(* IEC 61131-3 sources: plc-st-coding-agent/progress/evidence/v13_rescore_20261108b/candidates/custom_deepseek-v4pro, 35 files *)

(* ---- public-easy-01.st ---- *)
FUNCTION_BLOCK FB
VAR_INPUT
    bottleSensor: BOOL;
    cleaningConfirmButton: BOOL;
    fillingConfirmButton: BOOL;
    cappingConfirmButton: BOOL;
    packingConfirmButton: BOOL;
    finishedButton: BOOL;
END_VAR
VAR_OUTPUT
    Pump_Motor: BOOL;
    Filling_Valve: BOOL;
    Capping_Machine: BOOL;
    Packing_Machine: BOOL;
    Completion_Light: BOOL;
END_VAR
VAR
    step: INT := 0;
END_VAR

IF finishedButton THEN
    step := 0;
    Pump_Motor := FALSE;
    Filling_Valve := FALSE;
    Capping_Machine := FALSE;
    Packing_Machine := FALSE;
    Completion_Light := FALSE;
ELSE
    CASE step OF
        0:
            IF bottleSensor THEN
                step := 1;
                Pump_Motor := TRUE;
                Filling_Valve := FALSE;
                Capping_Machine := FALSE;
                Packing_Machine := FALSE;
                Completion_Light := FALSE;
            ELSE
                Pump_Motor := FALSE;
                Filling_Valve := FALSE;
                Capping_Machine := FALSE;
                Packing_Machine := FALSE;
                Completion_Light := FALSE;
            END_IF

        1:
            Pump_Motor := TRUE;
            Filling_Valve := FALSE;
            Capping_Machine := FALSE;
            Packing_Machine := FALSE;
            Completion_Light := FALSE;
            IF cleaningConfirmButton THEN
                step := 2;
                Filling_Valve := TRUE;
            END_IF

        2:
            Pump_Motor := TRUE;
            Filling_Valve := TRUE;
            Capping_Machine := FALSE;
            Packing_Machine := FALSE;
            Completion_Light := FALSE;
            IF fillingConfirmButton THEN
                step := 3;
                Capping_Machine := TRUE;
            END_IF

        3:
            Pump_Motor := TRUE;
            Filling_Valve := TRUE;
            Capping_Machine := TRUE;
            Packing_Machine := FALSE;
            Completion_Light := FALSE;
            IF cappingConfirmButton THEN
                step := 4;
                Packing_Machine := TRUE;
            END_IF

        4:
            Pump_Motor := TRUE;
            Filling_Valve := TRUE;
            Capping_Machine := TRUE;
            Packing_Machine := TRUE;
            Completion_Light := FALSE;
            IF packingConfirmButton THEN
                step := 5;
                Completion_Light := TRUE;
            END_IF

        5:
            Pump_Motor := TRUE;
            Filling_Valve := TRUE;
            Capping_Machine := TRUE;
            Packing_Machine := TRUE;
            Completion_Light := TRUE;

    ELSE
        step := 0;
        Pump_Motor := FALSE;
        Filling_Valve := FALSE;
        Capping_Machine := FALSE;
        Packing_Machine := FALSE;
        Completion_Light := FALSE;
    END_CASE
END_IF

END_FUNCTION_BLOCK

(* ---- public-easy-02.st ---- *)
FUNCTION_BLOCK FB
VAR_INPUT
    value : DWORD;
END_VAR
VAR_OUTPUT
    hasChanged : BOOL;
    hasRisingEdges : BOOL;
    risingBits : DWORD;
    noOfRisingBits : USINT;
    hasFallingEdges : BOOL;
    fallingBits : DWORD;
    noOfFallingBits : USINT;
END_VAR
VAR
    previousValue : DWORD := 0;
    bitIndex : INT;
END_VAR
    risingBits := value AND (NOT previousValue);
    fallingBits := (NOT value) AND previousValue;

    hasRisingEdges := risingBits <> 0;
    hasFallingEdges := fallingBits <> 0;
    hasChanged := hasRisingEdges OR hasFallingEdges;

    noOfRisingBits := 0;
    noOfFallingBits := 0;
    FOR bitIndex := 0 TO 31 DO
        IF (risingBits AND SHL(DWORD#1, bitIndex)) <> 0 THEN
            noOfRisingBits := noOfRisingBits + 1;
        END_IF;
        IF (fallingBits AND SHL(DWORD#1, bitIndex)) <> 0 THEN
            noOfFallingBits := noOfFallingBits + 1;
        END_IF;
    END_FOR;

    previousValue := value;
END_FUNCTION_BLOCK

(* ---- public-easy-03.st ---- *)
FUNCTION_BLOCK FB
VAR_INPUT
    Value : REAL;
    hiLevel : REAL;
    loLevel : REAL;
    hystWindow : REAL;
END_VAR
VAR_OUTPUT
    hiAlarm : BOOL;
    loAlarm : BOOL;
    error : BOOL;
    status : WORD;
END_VAR
VAR
END_VAR

error := FALSE;
status := 0;

IF loLevel >= hiLevel THEN
    error := TRUE;
    status := 16#8001;
ELSIF hystWindow >= (hiLevel - loLevel) THEN
    error := TRUE;
    status := 16#8002;
ELSE
    IF Value > hiLevel THEN
        hiAlarm := TRUE;
    ELSIF Value < (hiLevel - hystWindow) THEN
        hiAlarm := FALSE;
    END_IF;

    IF Value < loLevel THEN
        loAlarm := TRUE;
    ELSIF Value > (loLevel + hystWindow) THEN
        loAlarm := FALSE;
    END_IF;
END_IF;

END_FUNCTION_BLOCK

(* ---- public-easy-04.st ---- *)
FUNCTION_BLOCK FB
VAR_INPUT
    VISCOSITY_OK: BOOL;
    PASTE_E_STOP_NC: BOOL;
    DebounceTime: TIME;
    CycleTime: TIME;
END_VAR
VAR_OUTPUT
    VFD_RUN: BOOL;
    PUMP_MAINT_DUE: BOOL;
    PUMP_RUNTIME_ACC: LINT;
END_VAR
VAR
    DebounceAccum: LINT := 0;               (* Debounce accumulated time in ms *)
    AccumRuntime: LINT := 0;                (* Accumulated pump runtime in ms *)
    MaintDue: BOOL := FALSE;                (* Maintenance due latch *)
    DebounceTimeMs: LINT := 0;              (* DebounceTime in ms *)
    MAINT_THRESHOLD: LINT := 1800000000;    (* 500 hours in ms *)
END_VAR

(* Convert DebounceTime to milliseconds (CODESYS TIME_TO_LINT preserves ms value) *)
DebounceTimeMs := TIME_TO_LINT(DebounceTime);

(* Debounce logic with E-stop priority:
   - VISCOSITY_OK FALSE immediately clears debounce.
   - E-stop active clears only incomplete debounce, keeps completed condition.
   - Normal condition accumulates when signal is stable and E-stop is OK.
*)
IF NOT VISCOSITY_OK THEN
    DebounceAccum := 0;
ELSIF NOT PASTE_E_STOP_NC THEN
    IF DebounceAccum < DebounceTimeMs THEN
        DebounceAccum := 0;
    END_IF;
ELSE
    IF DebounceAccum < DebounceTimeMs THEN
        DebounceAccum := DebounceAccum + TIME_TO_LINT(CycleTime);
        IF DebounceAccum > DebounceTimeMs THEN
            DebounceAccum := DebounceTimeMs;
        END_IF;
    END_IF;
END_IF;

(* Run command requires E-stop OK, viscosity raw signal TRUE and debounced condition valid *)
VFD_RUN := PASTE_E_STOP_NC AND VISCOSITY_OK AND (DebounceAccum >= DebounceTimeMs);

(* Accumulate enabled runtime only while pump is running *)
IF VFD_RUN THEN
    AccumRuntime := AccumRuntime + TIME_TO_LINT(CycleTime);
END_IF;

(* Maintenance due latch when accumulated time reaches 500 hours (1,800,000,000 ms) *)
IF AccumRuntime >= MAINT_THRESHOLD THEN
    MaintDue := TRUE;
END_IF;

(* Map internal state to outputs *)
PUMP_RUNTIME_ACC := AccumRuntime;
PUMP_MAINT_DUE := MaintDue;

END_FUNCTION_BLOCK

(* ---- public-easy-05.st ---- *)
FUNCTION_BLOCK FB
VAR_INPUT
    Gap_Exceeded : BOOL;
    Weld_E_Stop_NC : BOOL;
    DebounceTime : TIME;
END_VAR
VAR_OUTPUT
    Operator_Alert : BOOL;
    Weld_Soft_Start_Active : BOOL;
END_VAR
VAR
    init_count : DINT := 0;
    debounce_count : DINT := 0;
    InitPeriods : DINT := 5;
    DebouncePeriods : DINT;
END_VAR

DebouncePeriods := TIME_TO_DINT(DebounceTime);
IF DebouncePeriods < 3 THEN
    DebouncePeriods := 3;
END_IF;

Weld_Soft_Start_Active := (init_count < InitPeriods);

IF init_count < InitPeriods THEN
    init_count := init_count + 1;
END_IF;

IF NOT Weld_E_Stop_NC THEN
    Operator_Alert := FALSE;
    debounce_count := 0;
ELSE
    IF Weld_Soft_Start_Active THEN
        Operator_Alert := FALSE;
        debounce_count := 0;
    ELSE
        IF Gap_Exceeded THEN
            IF debounce_count < DebouncePeriods THEN
                debounce_count := debounce_count + 1;
            END_IF;
            IF debounce_count >= DebouncePeriods THEN
                Operator_Alert := TRUE;
            ELSE
                Operator_Alert := FALSE;
            END_IF;
        ELSE
            debounce_count := 0;
            Operator_Alert := FALSE;
        END_IF;
    END_IF;
END_IF;

END_FUNCTION_BLOCK

(* ---- public-easy-06.st ---- *)
FUNCTION_BLOCK FB
VAR_INPUT
    DO_LOW : BOOL;
    AERATION_E_STOP_NC : BOOL;
END_VAR
VAR_OUTPUT
    BLOWER_RUN : BOOL;
    AERATION_BLOWER_CYCLE_COUNT : UINT;
END_VAR
VAR
    timer_count : UINT := 0;
    last_run : BOOL := FALSE;
    run_cmd : BOOL := FALSE;
    cycle_count : UINT := 0;
END_VAR

IF DO_LOW AND AERATION_E_STOP_NC THEN
    IF timer_count < 5 THEN
        timer_count := timer_count + 1;
    END_IF;
ELSE
    timer_count := 0;
END_IF;

run_cmd := DO_LOW AND AERATION_E_STOP_NC AND (timer_count >= 5);

IF run_cmd AND NOT last_run THEN
    cycle_count := cycle_count + 1;
END_IF;

BLOWER_RUN := run_cmd;
AERATION_BLOWER_CYCLE_COUNT := cycle_count;
last_run := run_cmd;

END_FUNCTION_BLOCK

(* ---- public-hard-01.st ---- *)
FUNCTION_BLOCK FB
VAR_INPUT
    estop : BOOL;
    opeMode : BOOL;
    valveAStart : BOOL;
    valveBStart : BOOL;
    valveCStart : BOOL;
    valveDStart : BOOL;
    mixMotorStart : BOOL;
    autoStart : BOOL;
    processMode : BOOL;
    levelSensor : INT;
    mixMotorComplete : BOOL;
END_VAR
VAR_OUTPUT
    valveARun : BOOL;
    valveBRun : BOOL;
    valveCRun : BOOL;
    valveDRun : BOOL;
    mixMotorRun : BOOL;
END_VAR
VAR
    manValveA : BOOL := FALSE;
    manValveB : BOOL := FALSE;
    manValveC : BOOL := FALSE;
    manValveD : BOOL := FALSE;
    manMixMotor : BOOL := FALSE;
    autoStep : INT := 0;
    autoValveA : BOOL := FALSE;
    autoValveB : BOOL := FALSE;
    autoValveC : BOOL := FALSE;
    autoValveD : BOOL := FALSE;
    autoMixMotor : BOOL := FALSE;
    lastValveAStart : BOOL := FALSE;
    lastValveBStart : BOOL := FALSE;
    lastValveCStart : BOOL := FALSE;
    lastValveDStart : BOOL := FALSE;
    lastMixMotorStart : BOOL := FALSE;
    lastAutoStart : BOOL := FALSE;
    lastMixMotorComplete : BOOL := FALSE;
    lastOpeMode : BOOL := FALSE;
    valveAStartRising : BOOL;
    valveBStartRising : BOOL;
    valveCStartRising : BOOL;
    valveDStartRising : BOOL;
    mixMotorStartRising : BOOL;
    autoStartRising : BOOL;
    mixMotorCompleteRising : BOOL;
END_VAR

// 计算所有输入信号的上升沿
valveAStartRising := valveAStart AND NOT lastValveAStart;
valveBStartRising := valveBStart AND NOT lastValveBStart;
valveCStartRising := valveCStart AND NOT lastValveCStart;
valveDStartRising := valveDStart AND NOT lastValveDStart;
mixMotorStartRising := mixMotorStart AND NOT lastMixMotorStart;
autoStartRising := autoStart AND NOT lastAutoStart;
mixMotorCompleteRising := mixMotorComplete AND NOT lastMixMotorComplete;

// 急停或模式切换时，复位所有内部状态（手动记忆和自动步序）
IF (estop = FALSE) OR (opeMode <> lastOpeMode) THEN
    manValveA := FALSE;
    manValveB := FALSE;
    manValveC := FALSE;
    manValveD := FALSE;
    manMixMotor := FALSE;
    autoStep := 0;
    autoValveA := FALSE;
    autoValveB := FALSE;
    autoValveC := FALSE;
    autoValveD := FALSE;
    autoMixMotor := FALSE;
END_IF;

// 根据急停和模式设置输出
IF estop = TRUE THEN
    IF opeMode = FALSE THEN
        // 手动模式：按钮上升沿翻转对应输出
        IF valveAStartRising THEN
            manValveA := NOT manValveA;
        END_IF;
        IF valveBStartRising THEN
            manValveB := NOT manValveB;
        END_IF;
        IF valveCStartRising THEN
            manValveC := NOT manValveC;
        END_IF;
        IF valveDStartRising THEN
            manValveD := NOT manValveD;
        END_IF;
        IF mixMotorStartRising THEN
            manMixMotor := NOT manMixMotor;
        END_IF;

        valveARun := manValveA;
        valveBRun := manValveB;
        valveCRun := manValveC;
        valveDRun := manValveD;
        mixMotorRun := manMixMotor;
    ELSE
        // 自动模式
        IF autoStartRising THEN
            autoStep := 1;  // 进入FILL_A
            autoValveA := TRUE;
            autoValveB := FALSE;
            autoValveC := FALSE;
            autoValveD := FALSE;
            autoMixMotor := FALSE;
        END_IF;

        CASE autoStep OF
            0: // 空闲
                autoValveA := FALSE;
                autoValveB := FALSE;
                autoValveC := FALSE;
                autoValveD := FALSE;
                autoMixMotor := FALSE;

            1: // 填充A
                autoValveA := TRUE;
                autoValveB := FALSE;
                autoValveC := FALSE;
                autoValveD := FALSE;
                autoMixMotor := FALSE;
                IF levelSensor >= 50 THEN
                    autoValveA := FALSE;
                    autoStep := 2;
                END_IF;

            2: // 填充B
                autoValveB := TRUE;
                autoValveA := FALSE;
                autoValveC := FALSE;
                autoValveD := FALSE;
                autoMixMotor := FALSE;
                IF levelSensor >= 80 THEN
                    autoValveB := FALSE;
                    IF processMode THEN
                        autoStep := 4; // 填充C
                    ELSE
                        autoStep := 3; // 混合
                    END_IF;
                END_IF;

            3: // 混合电机运行
                autoMixMotor := TRUE;
                autoValveA := FALSE;
                autoValveB := FALSE;
                autoValveC := FALSE;
                autoValveD := FALSE;
                IF mixMotorCompleteRising THEN
                    autoMixMotor := FALSE;
                    autoValveD := TRUE;
                    autoStep := 5; // 出料
                END_IF;

            4: // 填充C（仅processMode=TRUE）
                autoValveC := TRUE;
                autoValveA := FALSE;
                autoValveB := FALSE;
                autoValveD := FALSE;
                autoMixMotor := FALSE;
                IF levelSensor >= 100 THEN
                    autoValveC := FALSE;
                    autoStep := 3; // 混合
                END_IF;

            5: // 出料
                autoValveD := TRUE;
                autoValveA := FALSE;
                autoValveB := FALSE;
                autoValveC := FALSE;
                autoMixMotor := FALSE;
                // 等待新的autoStart上升沿，由外层处理

            ELSE
                // 非法状态，复位
                autoStep := 0;
                autoValveA := FALSE;
                autoValveB := FALSE;
                autoValveC := FALSE;
                autoValveD := FALSE;
                autoMixMotor := FALSE;
        END_CASE;

        valveARun := autoValveA;
        valveBRun := autoValveB;
        valveCRun := autoValveC;
        valveDRun := autoValveD;
        mixMotorRun := autoMixMotor;
    END_IF;
ELSE
    // 急停触发：所有输出停止
    valveARun := FALSE;
    valveBRun := FALSE;
    valveCRun := FALSE;
    valveDRun := FALSE;
    mixMotorRun := FALSE;
END_IF;

// 更新历史值
lastValveAStart := valveAStart;
lastValveBStart := valveBStart;
lastValveCStart := valveCStart;
lastValveDStart := valveDStart;
lastMixMotorStart := mixMotorStart;
lastAutoStart := autoStart;
lastMixMotorComplete := mixMotorComplete;
lastOpeMode := opeMode;

END_FUNCTION_BLOCK

(* ---- public-hard-02.st ---- *)
FUNCTION_BLOCK FB
VAR_INPUT
    processLength : USINT;
    sensor1 : BOOL;
    sensor2 : BOOL;
    sensor3 : BOOL;
    sensor4 : BOOL;
    sensor5 : BOOL;
    station1Start : BOOL;
    station2Complete : BOOL;
    station3Complete : BOOL;
    station4Complete : BOOL;
    processSequence : ARRAY[1..8] OF USINT;
END_VAR
VAR_OUTPUT
    conveyorLeft : BOOL;
    conveyorRight : BOOL;
END_VAR
VAR
    phase : USINT := 0;
    curStation : USINT := 1;
    idx : USINT := 1;
    dstStation : USINT := 0;
    station1StartPrev : BOOL := FALSE;
    station2CompletePrev : BOOL := FALSE;
    station3CompletePrev : BOOL := FALSE;
    station4CompletePrev : BOOL := FALSE;
    sensor2Prev : BOOL := FALSE;
    sensor3Prev : BOOL := FALSE;
    sensor4Prev : BOOL := FALSE;
    sensor5Prev : BOOL := FALSE;
    station1StartRising : BOOL;
    station2CompleteRising : BOOL;
    station3CompleteRising : BOOL;
    station4CompleteRising : BOOL;
    sensor2Rising : BOOL;
    sensor3Rising : BOOL;
    sensor4Rising : BOOL;
    sensor5Rising : BOOL;
END_VAR

    station1StartRising := station1Start AND NOT station1StartPrev;
    station2CompleteRising := station2Complete AND NOT station2CompletePrev;
    station3CompleteRising := station3Complete AND NOT station3CompletePrev;
    station4CompleteRising := station4Complete AND NOT station4CompletePrev;
    sensor2Rising := sensor2 AND NOT sensor2Prev;
    sensor3Rising := sensor3 AND NOT sensor3Prev;
    sensor4Rising := sensor4 AND NOT sensor4Prev;
    sensor5Rising := sensor5 AND NOT sensor5Prev;

    IF phase = 0 THEN
        IF station1StartRising AND sensor1 THEN
            curStation := 1;
            idx := 1;
            dstStation := processSequence[idx];
            phase := 1;
        END_IF;
    ELSIF phase = 1 THEN
        IF (dstStation = 2 AND sensor2Rising) OR
           (dstStation = 3 AND sensor3Rising) OR
           (dstStation = 4 AND sensor4Rising) OR
           (dstStation = 5 AND sensor5Rising) THEN
            curStation := dstStation;
            IF dstStation = 5 THEN
                phase := 0;
                idx := 0;
            ELSE
                phase := 2;
            END_IF;
        END_IF;
    ELSIF phase = 2 THEN
        IF (curStation = 2 AND station2CompleteRising) OR
           (curStation = 3 AND station3CompleteRising) OR
           (curStation = 4 AND station4CompleteRising) THEN
            idx := idx + 1;
            dstStation := processSequence[idx];
            phase := 1;
        END_IF;
    ELSE
        phase := 0;
    END_IF;

    IF phase = 1 THEN
        IF dstStation > curStation THEN
            conveyorRight := TRUE;
            conveyorLeft := FALSE;
        ELSIF dstStation < curStation THEN
            conveyorLeft := TRUE;
            conveyorRight := FALSE;
        ELSE
            conveyorLeft := FALSE;
            conveyorRight := FALSE;
        END_IF;
    ELSE
        conveyorLeft := FALSE;
        conveyorRight := FALSE;
    END_IF;

    station1StartPrev := station1Start;
    station2CompletePrev := station2Complete;
    station3CompletePrev := station3Complete;
    station4CompletePrev := station4Complete;
    sensor2Prev := sensor2;
    sensor3Prev := sensor3;
    sensor4Prev := sensor4;
    sensor5Prev := sensor5;

END_FUNCTION_BLOCK

(* ---- public-hard-03.st ---- *)
TYPE ST_Recipe :
STRUCT
    recipeID : INT;
    ingredientType : INT;
    ingredientRatio : REAL;
    productionTemperature : REAL;
END_STRUCT
END_TYPE

FUNCTION_BLOCK FB
VAR_INPUT
    addRecipe : BOOL;
    deleteRecipe : BOOL;
    modifyRecipe : BOOL;
    queryRecipe : BOOL;
    recipeIn : ST_Recipe;
END_VAR
VAR_OUTPUT
    recipeAdded : BOOL;
    recipeDeleted : BOOL;
    recipeModified : BOOL;
    recipeQueryResult : ST_Recipe;
    error : BOOL;
    status : WORD;
END_VAR
VAR_IN_OUT
    recipe : ARRAY[1..10] OF ST_Recipe;
END_VAR
VAR
    prevAddRecipe : BOOL := FALSE;
    prevDeleteRecipe : BOOL := FALSE;
    prevModifyRecipe : BOOL := FALSE;
    prevQueryRecipe : BOOL := FALSE;
    addRising : BOOL;
    deleteRising : BOOL;
    modifyRising : BOOL;
    queryRising : BOOL;
    i : INT;
    foundIndex : INT;
    found : BOOL;
    emptyIndex : INT;
    duplicate : BOOL;
END_VAR

// 默认输出复位
recipeAdded := FALSE;
recipeDeleted := FALSE;
recipeModified := FALSE;
error := FALSE;
status := 0;

// 计算上升沿
addRising := addRecipe AND NOT prevAddRecipe;
deleteRising := deleteRecipe AND NOT prevDeleteRecipe;
modifyRising := modifyRecipe AND NOT prevModifyRecipe;
queryRising := queryRecipe AND NOT prevQueryRecipe;

// 更新历史状态
prevAddRecipe := addRecipe;
prevDeleteRecipe := deleteRecipe;
prevModifyRecipe := modifyRecipe;
prevQueryRecipe := queryRecipe;

// 按优先级处理请求（假设同一时刻只有一个请求被触发）
IF addRising THEN
    // 检查重复
    duplicate := FALSE;
    FOR i := 1 TO 10 DO
        IF recipe[i].recipeID <> 0 AND recipe[i].recipeID = recipeIn.recipeID THEN
            duplicate := TRUE;
            EXIT;
        END_IF;
    END_FOR;

    IF duplicate THEN
        error := TRUE;
        status := 16#8002;
    ELSE
        // 查找第一个空槽
        emptyIndex := 0;
        FOR i := 1 TO 10 DO
            IF recipe[i].recipeID = 0 THEN
                emptyIndex := i;
                EXIT;
            END_IF;
        END_FOR;

        IF emptyIndex = 0 THEN
            error := TRUE;
            status := 16#8003;
        ELSE
            recipe[emptyIndex] := recipeIn;
            recipeAdded := TRUE;
        END_IF;
    END_IF;
ELSIF deleteRising THEN
    // 查找要删除的配方
    found := FALSE;
    FOR i := 1 TO 10 DO
        IF recipe[i].recipeID <> 0 AND recipe[i].recipeID = recipeIn.recipeID THEN
            found := TRUE;
            foundIndex := i;
            EXIT;
        END_IF;
    END_FOR;

    IF NOT found THEN
        error := TRUE;
        status := 16#8004;
    ELSE
        recipe[foundIndex].recipeID := 0;
        recipeDeleted := TRUE;
    END_IF;
ELSIF modifyRising THEN
    // 查找要修改的配方
    found := FALSE;
    FOR i := 1 TO 10 DO
        IF recipe[i].recipeID <> 0 AND recipe[i].recipeID = recipeIn.recipeID THEN
            found := TRUE;
            foundIndex := i;
            EXIT;
        END_IF;
    END_FOR;

    IF NOT found THEN
        error := TRUE;
        status := 16#8005;
    ELSE
        recipe[foundIndex] := recipeIn;
        recipeModified := TRUE;
    END_IF;
ELSIF queryRising THEN
    // 查找要查询的配方
    found := FALSE;
    FOR i := 1 TO 10 DO
        IF recipe[i].recipeID <> 0 AND recipe[i].recipeID = recipeIn.recipeID THEN
            found := TRUE;
            recipeQueryResult := recipe[i];
            EXIT;
        END_IF;
    END_FOR;

    IF NOT found THEN
        error := TRUE;
        status := 16#8001;
    END_IF;
END_IF;

END_FUNCTION_BLOCK

(* ---- public-hard-04.st ---- *)
FUNCTION_BLOCK FB
VAR_INPUT
    enqueue : BOOL;
    dequeue : BOOL;
    reset : BOOL;
    capacity : DINT;
END_VAR
VAR_OUTPUT
    elementCount : DINT;
    status : WORD;
END_VAR
VAR_IN_OUT
    item : DINT;
    buffer : ARRAY[1..4] OF DINT;
END_VAR
VAR
    head : DINT := 1;
    tail : DINT := 1;
    count : DINT := 0;
    lastEnq : BOOL := FALSE;
    lastDeq : BOOL := FALSE;
    enqRising : BOOL;
    deqRising : BOOL;
END_VAR

// 计算上升沿
enqRising := enqueue AND NOT lastEnq;
deqRising := dequeue AND NOT lastDeq;

// 更新历史值
lastEnq := enqueue;
lastDeq := dequeue;

// 复位优先
IF reset THEN
    count := 0;
    head := 1;
    tail := 1;
    status := 16#0000;
ELSE
    // 入队操作
    IF enqRising THEN
        IF count < capacity THEN
            buffer[tail] := item;
            tail := tail + 1;
            IF tail > capacity THEN
                tail := 1;
            END_IF
            count := count + 1;
            status := 16#0000;
        ELSE
            status := 16#8002; // 队列满，入队被拒绝
        END_IF
    // 出队操作
    ELSIF deqRising THEN
        IF count > 0 THEN
            item := buffer[head];
            head := head + 1;
            IF head > capacity THEN
                head := 1;
            END_IF
            count := count - 1;
            status := 16#0000;
        ELSE
            status := 16#8001; // 队列空，出队被拒绝
        END_IF
    ELSE
        status := 16#0000;
    END_IF
END_IF

// 更新输出元素个数
elementCount := count;

END_FUNCTION_BLOCK

(* ---- public-hard-05.st ---- *)
FUNCTION_BLOCK FB
VAR_INPUT
    ManualMode : BOOL;
    SingleStepMode : BOOL;
    SingleCycleMode : BOOL;
    ContinuousMode : BOOL;
    EmergencyStop : BOOL;
    Start : BOOL;
    DownButton : BOOL;
    UpButton : BOOL;
    LeftButton : BOOL;
    RightButton : BOOL;
    GripButton : BOOL;
    ReleaseButton : BOOL;
    DownLimitSwitch : BOOL;
    UpLimitSwitch : BOOL;
    LeftLimitSwitch : BOOL;
    RightLimitSwitch : BOOL;
    GripLimitSwitch : BOOL;
    ReleaseLimitSwitch : BOOL;
END_VAR
VAR_OUTPUT
    MoveDown : BOOL;
    MoveUp : BOOL;
    MoveLeft : BOOL;
    MoveRight : BOOL;
    ActivateGrip : BOOL;
    ActivateRelease : BOOL;
END_VAR
VAR
    StartRise : BOOL;
    StartPrev : BOOL;
    AutoModeActive : BOOL;
    PrevAutoModeActive : BOOL;
    StepIndex : INT := 1;
    WaitingForStart : BOOL := TRUE;
    ManMoveDown : BOOL;
    ManMoveUp : BOOL;
    ManMoveLeft : BOOL;
    ManMoveRight : BOOL;
    ManGrip : BOOL;
    ManRelease : BOOL;
    AutoMoveDown : BOOL;
    AutoMoveUp : BOOL;
    AutoMoveLeft : BOOL;
    AutoMoveRight : BOOL;
    AutoGrip : BOOL;
    AutoRelease : BOOL;
    ReqMoveDown : BOOL;
    ReqMoveUp : BOOL;
    ReqMoveLeft : BOOL;
    ReqMoveRight : BOOL;
    ReqGrip : BOOL;
    ReqRelease : BOOL;
    StepDone : BOOL;
END_VAR

StartRise := Start AND NOT StartPrev;
StartPrev := Start;

AutoModeActive := SingleStepMode OR SingleCycleMode OR ContinuousMode;

IF AutoModeActive AND NOT PrevAutoModeActive THEN
    StepIndex := 1;
    WaitingForStart := TRUE;
END_IF;
PrevAutoModeActive := AutoModeActive;

ManMoveDown := ManualMode AND DownButton AND NOT DownLimitSwitch;
ManMoveUp := ManualMode AND UpButton AND NOT UpLimitSwitch;
ManMoveLeft := ManualMode AND LeftButton AND NOT LeftLimitSwitch;
ManMoveRight := ManualMode AND RightButton AND NOT RightLimitSwitch;
ManGrip := ManualMode AND GripButton AND NOT GripLimitSwitch;
ManRelease := ManualMode AND ReleaseButton AND NOT ReleaseLimitSwitch;

IF EmergencyStop THEN
    IF AutoModeActive THEN
        IF WaitingForStart THEN
            IF StartRise THEN
                WaitingForStart := FALSE;
            END_IF;
        ELSE
            StepDone := FALSE;
            CASE StepIndex OF
                1: StepDone := DownLimitSwitch;
                2: StepDone := GripLimitSwitch;
                3: StepDone := UpLimitSwitch;
                4: StepDone := RightLimitSwitch;
                5: StepDone := DownLimitSwitch;
                6: StepDone := ReleaseLimitSwitch;
                7: StepDone := UpLimitSwitch;
                8: StepDone := LeftLimitSwitch;
            END_CASE;
            IF StepDone THEN
                IF SingleStepMode THEN
                    WaitingForStart := TRUE;
                    IF StepIndex >= 8 THEN
                        StepIndex := 1;
                    ELSE
                        StepIndex := StepIndex + 1;
                    END_IF;
                ELSIF SingleCycleMode THEN
                    IF StepIndex >= 8 THEN
                        StepIndex := 1;
                        WaitingForStart := TRUE;
                    ELSE
                        StepIndex := StepIndex + 1;
                    END_IF;
                ELSIF ContinuousMode THEN
                    IF StepIndex >= 8 THEN
                        StepIndex := 1;
                    ELSE
                        StepIndex := StepIndex + 1;
                    END_IF;
                END_IF;
            END_IF;
        END_IF;
    END_IF;
END_IF;

IF AutoModeActive AND NOT WaitingForStart THEN
    AutoMoveDown := (StepIndex = 1) OR (StepIndex = 5);
    AutoMoveUp := (StepIndex = 3) OR (StepIndex = 7);
    AutoMoveLeft := (StepIndex = 8);
    AutoMoveRight := (StepIndex = 4);
    AutoGrip := (StepIndex = 2);
    AutoRelease := (StepIndex = 6);
ELSE
    AutoMoveDown := FALSE;
    AutoMoveUp := FALSE;
    AutoMoveLeft := FALSE;
    AutoMoveRight := FALSE;
    AutoGrip := FALSE;
    AutoRelease := FALSE;
END_IF;

ReqMoveDown := ManMoveDown OR AutoMoveDown;
ReqMoveUp := ManMoveUp OR AutoMoveUp;
ReqMoveLeft := ManMoveLeft OR AutoMoveLeft;
ReqMoveRight := ManMoveRight OR AutoMoveRight;
ReqGrip := ManGrip OR AutoGrip;
ReqRelease := ManRelease OR AutoRelease;

MoveDown := ReqMoveDown AND NOT ReqMoveUp;
MoveUp := ReqMoveUp AND NOT ReqMoveDown;
MoveLeft := ReqMoveLeft AND NOT ReqMoveRight;
MoveRight := ReqMoveRight AND NOT ReqMoveLeft;
ActivateGrip := ReqGrip AND NOT ReqRelease;
ActivateRelease := ReqRelease AND NOT ReqGrip;

IF NOT EmergencyStop THEN
    MoveDown := FALSE;
    MoveUp := FALSE;
    MoveLeft := FALSE;
    MoveRight := FALSE;
    ActivateGrip := FALSE;
    ActivateRelease := FALSE;
END_IF;

END_FUNCTION_BLOCK

(* ---- public-hard-06.st ---- *)
FUNCTION_BLOCK FB
VAR_INPUT
    Mode : BOOL;
    ForwardButton : BOOL;
    ReverseButton : BOOL;
    SensorFeed : BOOL;
    SensorWash : BOOL;
    SensorWeight : BOOL;
    SensorFiring : BOOL;
    SensorOutput : BOOL;
    washComplete : BOOL;
    weightComplete : BOOL;
    weight : REAL;
    firingComplete : BOOL;
END_VAR
VAR_OUTPUT
    MotorForward : BOOL;
    MotorReverse : BOOL;
    kick : BOOL;
    CompletionLight : BOOL;
    firingTemp : REAL;
END_VAR
VAR
    state : INT := 0;
END_VAR

IF Mode THEN
    (* Automatic mode *)
    MotorReverse := FALSE;
    kick := FALSE;
    CompletionLight := FALSE;

    CASE state OF
        0: (* IDLE *)
            IF SensorFeed THEN
                state := 1;
            END_IF
        1: (* MOVING_TO_WASH *)
            IF SensorWash THEN
                state := 2;
            END_IF
        2: (* AT_WASH *)
            IF washComplete THEN
                state := 3;
            END_IF
        3: (* MOVING_TO_WEIGHT *)
            IF SensorWeight THEN
                state := 4;
            END_IF
        4: (* AT_WEIGHT *)
            IF weightComplete THEN
                IF weight >= 100.0 AND weight <= 200.0 THEN
                    firingTemp := 500.0 + (weight - 100.0) * (550.0 - 500.0) / (200.0 - 100.0);
                    state := 5;
                ELSE
                    kick := TRUE;
                    state := 9;
                END_IF
            END_IF
        5: (* MOVING_TO_FIRING *)
            IF SensorFiring THEN
                state := 6;
            END_IF
        6: (* AT_FIRING *)
            IF firingComplete THEN
                state := 7;
            END_IF
        7: (* MOVING_TO_OUTPUT *)
            IF SensorOutput THEN
                state := 8;
            END_IF
        8: (* AT_OUTPUT *)
            CompletionLight := TRUE;
            IF NOT SensorOutput THEN
                CompletionLight := FALSE;
                state := 0;
            END_IF
        9: (* REJECTING *)
            IF NOT SensorWeight THEN
                state := 0;
            END_IF
    END_CASE

    IF state = 1 OR state = 3 OR state = 5 OR state = 7 THEN
        MotorForward := TRUE;
    ELSE
        MotorForward := FALSE;
    END_IF

ELSE
    (* Manual mode *)
    MotorForward := ForwardButton AND NOT ReverseButton;
    MotorReverse := ReverseButton AND NOT ForwardButton;
    kick := FALSE;
    CompletionLight := FALSE;
    state := 0;
END_IF

END_FUNCTION_BLOCK

(* ---- public-medium-01.st ---- *)
TYPE ST_Pump :
STRUCT
    priority : INT;
    selection : BOOL;
    RunComd : BOOL;
END_STRUCT
END_TYPE

FUNCTION_BLOCK FB
VAR_INPUT
    mode : BOOL;
    start : BOOL;
    stop : BOOL;
END_VAR
VAR_IN_OUT
    pumpGroup : ARRAY[1..5] OF ST_Pump;
END_VAR
VAR
    prioArr : ARRAY[1..5] OF INT;
    idxArr : ARRAY[1..5] OF INT;
    i : INT;
    j : INT;
    tempPrio : INT;
    tempIdx : INT;
END_VAR

    IF stop OR NOT start THEN
        FOR i := 1 TO 5 DO
            pumpGroup[i].RunComd := FALSE;
        END_FOR
    ELSE
        IF NOT mode THEN
            FOR i := 1 TO 5 DO
                pumpGroup[i].RunComd := pumpGroup[i].selection;
            END_FOR
        ELSE
            FOR i := 1 TO 5 DO
                pumpGroup[i].RunComd := FALSE;
            END_FOR

            FOR i := 1 TO 5 DO
                prioArr[i] := pumpGroup[i].priority;
                idxArr[i] := i;
            END_FOR

            FOR i := 1 TO 4 DO
                FOR j := 1 TO 5 - i DO
                    IF (prioArr[j] < prioArr[j + 1]) OR
                       (prioArr[j] = prioArr[j + 1] AND (idxArr[j] > idxArr[j + 1])) THEN
                        tempPrio := prioArr[j];
                        prioArr[j] := prioArr[j + 1];
                        prioArr[j + 1] := tempPrio;
                        tempIdx := idxArr[j];
                        idxArr[j] := idxArr[j + 1];
                        idxArr[j + 1] := tempIdx;
                    END_IF
                END_FOR
            END_FOR

            FOR i := 1 TO 3 DO
                pumpGroup[idxArr[i]].RunComd := TRUE;
            END_FOR
        END_IF
    END_IF

END_FUNCTION_BLOCK

(* ---- public-medium-02.st ---- *)
TYPE ST_AnalogChannel :
STRUCT
    enable : BOOL;
    hiLIM : REAL;
    loLIM : REAL;
    bipolar : BOOL;
    measuringMode : INT;
    retVal : WORD;
    outputValue : REAL;
END_STRUCT
END_TYPE

FUNCTION_BLOCK FB
VAR_INPUT
    count : DINT;
END_VAR
VAR_IN_OUT
    analogValues : ARRAY[1..8] OF INT;
    channels : ARRAY[1..8] OF ST_AnalogChannel;
END_VAR
VAR
    i : INT;
    raw : INT;
    rawReal : REAL;
    mapped : REAL;
    rangeLow : REAL := -27648.0;
    rangeHigh : REAL := 27648.0;
    unipolarHigh : REAL := 27648.0;
    unipolarLow : REAL := 0.0;
    scaleSpan : REAL;
    rawSpan : REAL;
END_VAR

    FOR i := 1 TO 8 DO
        IF i > count THEN
            EXIT;
        END_IF;

        IF channels[i].enable THEN
            IF (channels[i].measuringMode = 0) OR
               (channels[i].measuringMode = 1) OR
               (channels[i].measuringMode = 2) THEN

                IF channels[i].hiLIM > channels[i].loLIM THEN
                    raw := analogValues[i];
                    rawReal := INT_TO_REAL(raw);

                    CASE channels[i].measuringMode OF
                        0:
                            IF channels[i].bipolar THEN
                                rawSpan := rangeHigh - rangeLow;  (* 55296.0 *)
                                scaleSpan := channels[i].hiLIM - channels[i].loLIM;
                                mapped := channels[i].loLIM +
                                          (rawReal - rangeLow) / rawSpan * scaleSpan;
                            ELSE
                                rawSpan := unipolarHigh - unipolarLow; (* 27648.0 *)
                                scaleSpan := channels[i].hiLIM - channels[i].loLIM;
                                mapped := channels[i].loLIM +
                                          (rawReal - unipolarLow) / rawSpan * scaleSpan;
                            END_IF;

                        1:
                            mapped := rawReal / 10.0;

                        2:
                            mapped := rawReal / 100.0;
                    ELSE
                        mapped := 0.0; (* should never be reached *)
                    END_CASE;

                    channels[i].outputValue := mapped;
                    channels[i].retVal := 0;
                ELSE
                    channels[i].retVal := 16#8002;
                    (* outputValue unchanged *)
                END_IF;

            ELSE
                channels[i].retVal := 16#8001;
                (* outputValue unchanged *)
            END_IF;

        (* enable = FALSE: nothing is written to retVal or outputValue *)
        END_IF;
    END_FOR;

END_FUNCTION_BLOCK

(* ---- public-medium-03.st ---- *)
FUNCTION_BLOCK FB
VAR_INPUT
    cyclicExecution : BOOL;
    trigger : BOOL;
    value : LREAL;
    windowSize : INT;
    reset : BOOL;
END_VAR
VAR_OUTPUT
    average : LREAL;
    windowSizeReached : BOOL;
    error : BOOL;
    status : WORD;
END_VAR
VAR
    buffer : ARRAY[0..99] OF LREAL;
    inIdx : INT := 0;
    outIdx : INT := 0;
    count : INT := 0;
    sum : LREAL := 0.0;
    lastTrigger : BOOL := FALSE;
    shouldRead : BOOL;
    oldest : LREAL;
END_VAR

IF reset THEN
    // 复位：清除所有数据状态
    count := 0;
    sum := 0.0;
    inIdx := 0;
    outIdx := 0;
    average := 0.0;
    windowSizeReached := FALSE;
    // 检查窗口尺寸并设置错误状态
    IF windowSize < 1 OR windowSize > 100 THEN
        error := TRUE;
        status := 16#8200;
    ELSE
        error := FALSE;
        status := 16#0000;
    END_IF;
    // 更新触发边沿记忆
    lastTrigger := trigger;
ELSE
    // 检查窗口尺寸有效性
    IF windowSize < 1 OR windowSize > 100 THEN
        error := TRUE;
        status := 16#8200;
        average := 0.0;
        windowSizeReached := FALSE;
        lastTrigger := trigger;
    ELSE
        error := FALSE;
        status := 16#0000;

        // 调整缓冲区大小：如果当前样本数大于窗口尺寸，移除最旧的样本
        WHILE count > windowSize DO
            oldest := buffer[outIdx];
            sum := sum - oldest;
            outIdx := outIdx + 1;
            IF outIdx >= 100 THEN
                outIdx := 0;
            END_IF;
            count := count - 1;
        END_WHILE;

        // 确定是否应读取新值
        shouldRead := cyclicExecution OR (trigger AND NOT lastTrigger);

        // 更新触发边沿记忆
        lastTrigger := trigger;

        IF shouldRead THEN
            // 写入新值到缓冲区
            buffer[inIdx] := value;
            inIdx := inIdx + 1;
            IF inIdx >= 100 THEN
                inIdx := 0;
            END_IF;

            IF count = windowSize THEN
                // 缓冲区已满：移除最旧样本
                oldest := buffer[outIdx];
                sum := sum - oldest;
                outIdx := outIdx + 1;
                IF outIdx >= 100 THEN
                    outIdx := 0;
                END_IF;
                // count 保持不变
            ELSE
                // 缓冲区未满：增加样本计数
                count := count + 1;
            END_IF;

            // 更新总和
            sum := sum + value;
        END_IF;

        // 计算移动平均
        IF count > 0 THEN
            average := sum / count;
        ELSE
            average := 0.0;
        END_IF;

        // 窗口是否已满
        windowSizeReached := (count >= windowSize);
    END_IF;
END_IF;

END_FUNCTION_BLOCK

(* ---- public-medium-04.st ---- *)
FUNCTION_BLOCK FB
VAR_INPUT
    TemperatureSensorInput : REAL;
    SetTemperature : REAL;
END_VAR
VAR_OUTPUT
    CurrentTemperature : REAL;
    SetTempDisplay : REAL;
    HeaterStatus : BOOL;
    OverheatProtection : BOOL;
    HeaterOutput : BOOL;
END_VAR
VAR
    sensor_fault : BOOL;
    heater_on_counter : INT := 0;
    protection_counter : INT := 0;
    protection_active : BOOL := FALSE;
END_VAR

    CurrentTemperature := TemperatureSensorInput;
    SetTempDisplay := SetTemperature;

    sensor_fault := (TemperatureSensorInput < 0.0) OR (TemperatureSensorInput > 100.0);

    IF protection_active THEN
        HeaterOutput := FALSE;
        HeaterStatus := FALSE;
        OverheatProtection := TRUE;
        heater_on_counter := 0;

        protection_counter := protection_counter + 1;
        IF protection_counter >= 3 THEN
            protection_active := FALSE;
            OverheatProtection := FALSE;
            protection_counter := 0;
        END_IF;
    ELSE
        OverheatProtection := FALSE;

        IF sensor_fault THEN
            HeaterOutput := FALSE;
            heater_on_counter := 0;
        ELSIF TemperatureSensorInput < SetTemperature THEN
            HeaterOutput := TRUE;
            heater_on_counter := heater_on_counter + 1;

            IF heater_on_counter >= 5 THEN
                protection_active := TRUE;
                OverheatProtection := TRUE;
                HeaterOutput := FALSE;
                heater_on_counter := 0;
                protection_counter := 0;
            END_IF;
        ELSE
            HeaterOutput := FALSE;
            heater_on_counter := 0;
        END_IF;

        HeaterStatus := HeaterOutput;
    END_IF;

END_FUNCTION_BLOCK

(* ---- public-medium-05.st ---- *)
FUNCTION_BLOCK FB
VAR_INPUT
    Mode : BOOL;
    ForwardButton : BOOL;
    ReverseButton : BOOL;
    SensorA : BOOL;
    SensorB : BOOL;
    SensorC : BOOL;
    ButtonA : BOOL;
    ButtonB : BOOL;
    ButtonC : BOOL;
END_VAR
VAR_OUTPUT
    MotorForward : BOOL;
    MotorReverse : BOOL;
    CompletionLight : BOOL;
END_VAR
VAR
    step : INT := 0;
    btnA_prev : BOOL := FALSE;
    btnB_prev : BOOL := FALSE;
    btnC_prev : BOOL := FALSE;
    mode_prev : BOOL := FALSE;
    btnA_rise : BOOL;
    btnB_rise : BOOL;
    btnC_rise : BOOL;
    mode_fall : BOOL;
    forward_req : BOOL := FALSE;
    completion_trig : BOOL := FALSE;
END_VAR

// Edge detection
btnA_rise := ButtonA AND NOT btnA_prev;
btnB_rise := ButtonB AND NOT btnB_prev;
btnC_rise := ButtonC AND NOT btnC_prev;
mode_fall := mode_prev AND NOT Mode;

// Update history
btnA_prev := ButtonA;
btnB_prev := ButtonB;
btnC_prev := ButtonC;
mode_prev := Mode;

// Clear automatic process on falling edge to manual
IF mode_fall THEN
    step := 0;
    forward_req := FALSE;
    completion_trig := FALSE;
END_IF;

IF Mode THEN
    // Automatic mode
    CASE step OF
        0:
            forward_req := FALSE;
            completion_trig := FALSE;
            IF SensorA AND btnA_rise THEN
                step := 1;
                forward_req := TRUE;
            END_IF;
        1:
            forward_req := TRUE;
            completion_trig := FALSE;
            IF SensorB THEN
                step := 2;
                forward_req := FALSE;
            END_IF;
        2:
            forward_req := FALSE;
            completion_trig := FALSE;
            IF SensorB AND btnB_rise THEN
                step := 3;
                forward_req := TRUE;
            END_IF;
        3:
            forward_req := TRUE;
            completion_trig := FALSE;
            IF SensorC THEN
                step := 4;
                forward_req := FALSE;
            END_IF;
        4:
            forward_req := FALSE;
            IF SensorC AND btnC_rise THEN
                completion_trig := TRUE;
            END_IF;
            IF NOT SensorC THEN
                completion_trig := FALSE;
                step := 0;
            END_IF;
    END_CASE;

    MotorForward := forward_req;
    MotorReverse := FALSE;
ELSE
    // Manual mode
    MotorForward := ForwardButton AND NOT ReverseButton;
    MotorReverse := ReverseButton AND NOT ForwardButton;
END_IF;

CompletionLight := Mode AND SensorC AND completion_trig;

END_FUNCTION_BLOCK

(* ---- public-medium-06.st ---- *)
FUNCTION_BLOCK FB
VAR_INPUT
    THICKNESS_FAULT: BOOL;
    THICKNESS_SIGNAL_VALID: BOOL;
    CUTTING_RUN: BOOL;
    FaultTimestamp: DINT;
    CycleTime: TIME;
END_VAR
VAR_OUTPUT
    THICKNESS_ALARM: BOOL := FALSE;
    Slab_Fault_Counter: UINT := 0;
    Slab_Runtime_Accumulator: LINT := 0;
    Slab_Fault_History: ARRAY[0..4] OF DINT := [0,0,0,0,0];
END_VAR
VAR
    faultPrev: BOOL := FALSE;
    alarmHoldTimer: TIME := T#0ms;
    i: INT;
END_VAR

IF NOT THICKNESS_SIGNAL_VALID THEN
    THICKNESS_ALARM := FALSE;
    alarmHoldTimer := T#0ms;
    faultPrev := FALSE;
ELSE
    IF THICKNESS_FAULT AND NOT faultPrev THEN
        Slab_Fault_Counter := Slab_Fault_Counter + 1;
        i := 4;
        WHILE i >= 1 DO
            Slab_Fault_History[i] := Slab_Fault_History[i-1];
            i := i - 1;
        END_WHILE;
        Slab_Fault_History[0] := FaultTimestamp;
    END_IF;

    IF THICKNESS_FAULT THEN
        THICKNESS_ALARM := TRUE;
        alarmHoldTimer := T#0ms;
    ELSE
        IF THICKNESS_ALARM THEN
            alarmHoldTimer := alarmHoldTimer + CycleTime;
            IF alarmHoldTimer >= T#500ms THEN
                THICKNESS_ALARM := FALSE;
                alarmHoldTimer := T#0ms;
            ELSE
                THICKNESS_ALARM := TRUE;
            END_IF;
        ELSE
            THICKNESS_ALARM := FALSE;
            alarmHoldTimer := T#0ms;
        END_IF;
    END_IF;

    IF CUTTING_RUN AND NOT THICKNESS_FAULT THEN
        Slab_Runtime_Accumulator := Slab_Runtime_Accumulator + TIME_TO_LINT(CycleTime);
    END_IF;

    faultPrev := THICKNESS_FAULT;
END_IF;

END_FUNCTION_BLOCK

(* ---- public-medium-07.st ---- *)
FUNCTION_BLOCK FB
VAR_INPUT
    OCCUPANCY_DETECTED: BOOL;
    ENERGY_SAVING_MODE: BOOL;
    HVAC_MODE_SELECTOR: INT;
END_VAR
VAR_OUTPUT
    SUPPLY_FAN_RUN: BOOL;
    TEMP_SETPOINT_ADJUST: INT;
END_VAR
VAR
    fan_delay_count: INT := 0;
END_VAR

(* Fan start delay logic - valid modes are 0(Auto),1(Comfort),2(Economy); Night(3) or invalid stop fan *)
IF OCCUPANCY_DETECTED AND (HVAC_MODE_SELECTOR >= 0) AND (HVAC_MODE_SELECTOR <= 2) THEN
    IF fan_delay_count < 30 THEN
        fan_delay_count := fan_delay_count + 1;
    END_IF;
    IF fan_delay_count >= 30 THEN
        SUPPLY_FAN_RUN := TRUE;
    ELSE
        SUPPLY_FAN_RUN := FALSE;
    END_IF;
ELSE
    fan_delay_count := 0;
    SUPPLY_FAN_RUN := FALSE;
END_IF;

(* Temperature setpoint adjustment *)
CASE HVAC_MODE_SELECTOR OF
    0: (* Auto *)
        IF OCCUPANCY_DETECTED THEN
            TEMP_SETPOINT_ADJUST := 0;
        ELSE
            IF ENERGY_SAVING_MODE THEN
                TEMP_SETPOINT_ADJUST := 3;
            ELSE
                TEMP_SETPOINT_ADJUST := 2;
            END_IF;
        END_IF;
    1: (* Comfort *)
        IF OCCUPANCY_DETECTED THEN
            TEMP_SETPOINT_ADJUST := 0;
        ELSE
            TEMP_SETPOINT_ADJUST := 1;
        END_IF;
    2: (* Economy *)
        IF OCCUPANCY_DETECTED THEN
            TEMP_SETPOINT_ADJUST := 0;
        ELSE
            TEMP_SETPOINT_ADJUST := 4;
        END_IF;
    3: (* Night *)
        TEMP_SETPOINT_ADJUST := 4;
    ELSE
        TEMP_SETPOINT_ADJUST := 0; (* invalid mode safe side *)
END_CASE;

END_FUNCTION_BLOCK

(* ---- public-medium-08.st ---- *)
FUNCTION_BLOCK FB
VAR_INPUT
    ipText : STRING(254);
END_VAR
VAR_OUTPUT
    ipValue : UDINT;
END_VAR
VAR
    ok : BOOL := FALSE;
    segCount : INT := 0;
    segLen : INT;
    segVal : UDINT;
    segIndex : INT;
    segVals : ARRAY[1..4] OF UDINT;
    textLen : INT;
    i : INT;
    ch : STRING(1);
END_VAR

// 初始化
ok := TRUE;
ipValue := 0;
segCount := 0;
segIndex := 1;
segLen := 0;
segVal := 0;
textLen := LEN(ipText);

FOR i := 1 TO textLen DO
    ch := MID(ipText, i, 1);
    IF ch = '.' THEN
        // 点：结束当前段
        IF segLen = 0 THEN
            ok := FALSE;
            EXIT;
        END_IF;
        IF segVal > 255 THEN
            ok := FALSE;
            EXIT;
        END_IF;
        IF segIndex > 4 THEN
            ok := FALSE;
            EXIT;
        END_IF;
        segVals[segIndex] := segVal;
        segIndex := segIndex + 1;
        // 重置当前段
        segVal := 0;
        segLen := 0;
    ELSIF ch = '0' THEN
        segVal := segVal * 10 + 0;
        segLen := segLen + 1;
    ELSIF ch = '1' THEN
        segVal := segVal * 10 + 1;
        segLen := segLen + 1;
    ELSIF ch = '2' THEN
        segVal := segVal * 10 + 2;
        segLen := segLen + 1;
    ELSIF ch = '3' THEN
        segVal := segVal * 10 + 3;
        segLen := segLen + 1;
    ELSIF ch = '4' THEN
        segVal := segVal * 10 + 4;
        segLen := segLen + 1;
    ELSIF ch = '5' THEN
        segVal := segVal * 10 + 5;
        segLen := segLen + 1;
    ELSIF ch = '6' THEN
        segVal := segVal * 10 + 6;
        segLen := segLen + 1;
    ELSIF ch = '7' THEN
        segVal := segVal * 10 + 7;
        segLen := segLen + 1;
    ELSIF ch = '8' THEN
        segVal := segVal * 10 + 8;
        segLen := segLen + 1;
    ELSIF ch = '9' THEN
        segVal := segVal * 10 + 9;
        segLen := segLen + 1;
    ELSE
        ok := FALSE;
        EXIT;
    END_IF;
END_FOR;

// 处理最后一个段
IF ok THEN
    IF segLen = 0 THEN
        ok := FALSE;
    ELSIF segVal > 255 THEN
        ok := FALSE;
    ELSIF segIndex > 4 THEN
        ok := FALSE;
    ELSE
        segVals[segIndex] := segVal;
        segIndex := segIndex + 1;
    END_IF;
END_IF;

// 最终判断
IF ok AND (segIndex - 1 = 4) THEN
    segCount := 4;
    ipValue := SHL(segVals[1], 24) OR SHL(segVals[2], 16) OR SHL(segVals[3], 8) OR segVals[4];
ELSE
    ok := FALSE;
    segCount := 0;
    ipValue := 0;
END_IF;

END_FUNCTION_BLOCK

(* ---- self-easy-01.st ---- *)
FUNCTION_BLOCK FB
VAR_INPUT
    enable : BOOL;
    values : ARRAY[1..8] OF INT;
    count : INT;
    avgEnable : BOOL;
END_VAR
VAR_OUTPUT
    avgOut : REAL;
END_VAR
VAR
    lastAvg : REAL := 0.0;
    actualCount : INT := 0;
    sum : DINT := 0;
    idx : INT := 0;
END_VAR

IF enable AND avgEnable THEN
    IF count <= 0 THEN
        actualCount := 0;
    ELSIF count > 8 THEN
        actualCount := 8;
    ELSE
        actualCount := count;
    END_IF;

    IF actualCount > 0 THEN
        sum := 0;
        FOR idx := 1 TO actualCount BY 1 DO
            sum := sum + INT_TO_DINT(values[idx]);
        END_FOR;
        lastAvg := DINT_TO_REAL(sum) / INT_TO_REAL(actualCount);
    END_IF;
END_IF;

avgOut := lastAvg;

END_FUNCTION_BLOCK

(* ---- self-easy-02.st ---- *)
FUNCTION_BLOCK FB
VAR_INPUT
    tankLevel : REAL;
    outletFlow : REAL;
    inletPermit : BOOL;
    resetBtn : BOOL;
END_VAR
VAR_OUTPUT
    pumpRun : BOOL;
    alarmHigh : BOOL;
    alarmLow : BOOL;
    outletValveOpen : BOOL;
END_VAR
VAR
    resetBtnPrev : BOOL;
    resetRising : BOOL;
    alarmHighState : BOOL;
    alarmLowState : BOOL;
END_VAR

resetRising := resetBtn AND NOT resetBtnPrev;

IF tankLevel >= 85.0 THEN
    alarmHighState := TRUE;
ELSIF resetRising THEN
    alarmHighState := FALSE;
END_IF

IF tankLevel <= 15.0 THEN
    alarmLowState := TRUE;
ELSIF resetRising THEN
    alarmLowState := FALSE;
END_IF

pumpRun := (tankLevel >= 15.0 AND tankLevel < 85.0) AND inletPermit AND NOT alarmHighState AND NOT alarmLowState;
outletValveOpen := (tankLevel >= 15.0 AND tankLevel < 85.0) AND inletPermit AND NOT alarmHighState AND NOT alarmLowState;

alarmHigh := alarmHighState;
alarmLow := alarmLowState;

resetBtnPrev := resetBtn;

END_FUNCTION_BLOCK

(* ---- self-hard-01.st ---- *)
FUNCTION_BLOCK FB
VAR_INPUT
    flowLow : BOOL;
    ackBtn : BOOL;
    sensorOK : BOOL;
END_VAR
VAR_OUTPUT
    alarmActive : BOOL;
    alarmAcked : BOOL;
    highHigh : BOOL;
END_VAR
VAR
    ackBtnPrev : BOOL := FALSE;
    ackRising : BOOL;
END_VAR

ackRising := ackBtn AND NOT ackBtnPrev;
ackBtnPrev := ackBtn;

highHigh := NOT sensorOK;

IF flowLow THEN
    IF ackRising THEN
        alarmActive := TRUE;
        alarmAcked := TRUE;
    ELSE
        alarmActive := TRUE;
        IF alarmAcked THEN
            alarmAcked := TRUE;
        ELSE
            alarmAcked := FALSE;
        END_IF
    END_IF
ELSE
    IF alarmActive THEN
        IF alarmAcked THEN
            alarmActive := FALSE;
            alarmAcked := FALSE;
        ELSE
            IF ackRising THEN
                alarmActive := FALSE;
                alarmAcked := FALSE;
            ELSE
                alarmActive := TRUE;
                alarmAcked := FALSE;
            END_IF
        END_IF
    ELSE
        alarmActive := FALSE;
        alarmAcked := FALSE;
    END_IF
END_IF

END_FUNCTION_BLOCK

(* ---- self-hard-02.st ---- *)
FUNCTION_BLOCK FB
VAR_INPUT
    startBtn : BOOL;
    abortBtn : BOOL;
    setpoint : REAL;
    pv : REAL;
    maxDuration : INT;
END_VAR
VAR_OUTPUT
    elapsed : INT;
    phase : INT;
    timeout : BOOL;
END_VAR
VAR
    lastStart : BOOL;
    startRising : BOOL;
END_VAR

    startRising := startBtn AND NOT lastStart;
    lastStart := startBtn;

    IF startRising THEN
        phase := 1;
        elapsed := 0;
        timeout := FALSE;
    ELSE
        IF abortBtn THEN
            phase := 9;
        ELSE
            IF phase = 1 OR phase = 2 THEN
                elapsed := elapsed + 1;
                IF elapsed >= maxDuration THEN
                    timeout := TRUE;
                    phase := 3;
                ELSE
                    IF phase = 1 THEN
                        IF pv >= setpoint THEN
                            phase := 2;
                        END_IF;
                    END_IF;
                END_IF;
            END_IF;
        END_IF;
    END_IF;

END_FUNCTION_BLOCK

(* ---- self-hard-03.st ---- *)
FUNCTION_BLOCK FB
VAR_INPUT
    pushEn : BOOL;
    pushItem : INT;
    popEn : BOOL;
END_VAR
VAR_IN_OUT
    fifo : ARRAY[1..8] OF INT;
END_VAR
VAR_OUTPUT
    count : INT;
    full : BOOL;
    empty : BOOL;
    head : INT;
END_VAR
VAR
    pushEn_prev : BOOL := FALSE;
    popEn_prev : BOOL := FALSE;
    pushRising : BOOL;
    popRising : BOOL;
    currentCount : INT := 0;
    i : INT;
END_VAR

pushRising := pushEn AND NOT pushEn_prev;
popRising := popEn AND NOT popEn_prev;

IF popRising AND (currentCount > 0) THEN
    IF currentCount > 1 THEN
        FOR i := 1 TO currentCount - 1 DO
            fifo[i] := fifo[i + 1];
        END_FOR;
    END_IF;
    fifo[currentCount] := 0;
    currentCount := currentCount - 1;
END_IF;

IF pushRising AND (currentCount < 8) THEN
    currentCount := currentCount + 1;
    fifo[currentCount] := pushItem;
END_IF;

pushEn_prev := pushEn;
popEn_prev := popEn;

count := currentCount;
full := (currentCount = 8);
empty := (currentCount = 0);

IF currentCount > 0 THEN
    head := fifo[1];
ELSE
    head := 0;
END_IF;

END_FUNCTION_BLOCK

(* ---- self-hard-04.st ---- *)
FUNCTION_BLOCK FB
VAR_INPUT
    demand : INT;
    runHours : ARRAY[1..5] OF LINT;
    rotated : BOOL;
END_VAR
VAR_OUTPUT
    leadPump : INT;
    lagPump : INT;
    runningCount : INT;
END_VAR
VAR
    orderedPumps : ARRAY[1..5] OF INT;
    initialized : BOOL := FALSE;
    tmpDemand : INT;
    tmpPump : INT;
    idx1 : INT;
    idx2 : INT;
END_VAR

tmpDemand := demand;
IF tmpDemand < 0 THEN
    tmpDemand := 0;
ELSIF tmpDemand > 5 THEN
    tmpDemand := 5;
END_IF

IF NOT initialized THEN
    FOR idx1 := 1 TO 5 DO
        orderedPumps[idx1] := idx1;
    END_FOR
    FOR idx1 := 1 TO 4 DO
        FOR idx2 := 1 TO 5 - idx1 DO
            IF runHours[orderedPumps[idx2]] > runHours[orderedPumps[idx2 + 1]] THEN
                tmpPump := orderedPumps[idx2];
                orderedPumps[idx2] := orderedPumps[idx2 + 1];
                orderedPumps[idx2 + 1] := tmpPump;
            END_IF
        END_FOR
    END_FOR
    initialized := TRUE;
END_IF

IF rotated THEN
    IF runHours[orderedPumps[2]] < (runHours[orderedPumps[1]] - 50) THEN
        tmpPump := orderedPumps[1];
        orderedPumps[1] := orderedPumps[2];
        orderedPumps[2] := tmpPump;
    END_IF
END_IF

IF tmpDemand = 0 THEN
    leadPump := 0;
    lagPump := 0;
    runningCount := 0;
ELSE
    leadPump := orderedPumps[1];
    runningCount := tmpDemand;
    IF tmpDemand >= 2 THEN
        lagPump := orderedPumps[2];
    ELSE
        lagPump := 0;
    END_IF
END_IF

END_FUNCTION_BLOCK

(* ---- self-hard-05.st ---- *)
FUNCTION_BLOCK FB
VAR_INPUT
    runRequest : BOOL;
    flameOK : BOOL;
    o2Valid : BOOL;
    o2PV : REAL;
    baseAir : REAL;
    resetBtn : BOOL;
END_VAR
VAR_OUTPUT
    fuelPermit : BOOL;
    trimEnable : BOOL;
    airTrim : REAL;
    airCommand : REAL;
    tripLatched : BOOL;
    o2Fault : BOOL;
END_VAR
VAR
    resetPrev : BOOL := FALSE;
    resRising : BOOL;
    tripState : BOOL := FALSE;
    trimRaw : REAL;
    airCmdRaw : REAL;
END_VAR

resRising := resetBtn AND NOT resetPrev;

IF runRequest AND NOT flameOK THEN
    tripState := TRUE;
ELSE
    IF resRising AND NOT runRequest AND NOT flameOK THEN
        tripState := FALSE;
    END_IF;
END_IF;

resetPrev := resetBtn;

tripLatched := tripState;

o2Fault := (NOT o2Valid) OR (o2PV < 0.0) OR (o2PV > 21.0);

fuelPermit := runRequest AND flameOK AND NOT tripState;

trimEnable := fuelPermit AND NOT o2Fault;

IF trimEnable THEN
    trimRaw := 2.0 * (2.0 - o2PV);
    IF trimRaw > 10.0 THEN
        trimRaw := 10.0;
    ELSIF trimRaw < -10.0 THEN
        trimRaw := -10.0;
    END_IF;
    airTrim := trimRaw;
ELSE
    airTrim := 0.0;
END_IF;

airCmdRaw := baseAir + airTrim;
IF airCmdRaw > 100.0 THEN
    airCmdRaw := 100.0;
ELSIF airCmdRaw < 0.0 THEN
    airCmdRaw := 0.0;
END_IF;

IF NOT fuelPermit THEN
    airCmdRaw := 0.0;
END_IF;

airCommand := airCmdRaw;

END_FUNCTION_BLOCK

(* ---- self-hard-06.st ---- *)
FUNCTION_BLOCK FB
VAR_INPUT
    runRequest : BOOL;
    pressure : REAL;
    pressureValid : BOOL;
    fuelFlow : REAL;
    steamFlow : REAL;
    outletCmd : INT;
    outletFeedback : INT;
    resetBtn : BOOL;
END_VAR
VAR_OUTPUT
    tripLatched : BOOL;
    fuelPermit : BOOL;
    currentCauseMask : WORD;
    latchedCauseMask : WORD;
    diagnosticActive : BOOL;
END_VAR
VAR
    resetBtnPrev : BOOL := FALSE;
    resetRising : BOOL;
    valveStuckCounter : INT := 0;
    tripCondition : BOOL;
    resetCondition : BOOL;
    bit1Active : BOOL;
    bit2Active : BOOL;
    stuckCond : BOOL;
END_VAR

// 卡滞条件判断，连续满足时计数
stuckCond := runRequest AND pressureValid AND (pressure >= 4500.0)
             AND (outletCmd >= 50) AND (outletFeedback <= 10);

IF stuckCond THEN
    valveStuckCounter := valveStuckCounter + 1;
ELSE
    valveStuckCounter := 0;
END_IF;

// 本周期诊断线索掩码计算
IF NOT runRequest THEN
    currentCauseMask := 0;
ELSIF NOT pressureValid THEN
    currentCauseMask := 16#0001; // bit0: 变送器失效
ELSE
    IF pressure >= 4500.0 THEN
        bit1Active := (valveStuckCounter >= 3);
        bit2Active := (fuelFlow >= 4.0) AND (steamFlow <= 10.0);
        IF bit1Active OR bit2Active THEN
            currentCauseMask := 0;
            IF bit1Active THEN
                currentCauseMask := currentCauseMask OR 16#0002; // bit1: 减温减压阀卡滞
            END_IF;
            IF bit2Active THEN
                currentCauseMask := currentCauseMask OR 16#0004; // bit2: 燃烧过剩
            END_IF;
        ELSE
            currentCauseMask := 16#0008; // bit3: 未定位
        END_IF;
    ELSE
        currentCauseMask := 0;
    END_IF;
END_IF;

// 复位按钮上升沿检测
resetRising := resetBtn AND NOT resetBtnPrev;

// 复位条件
resetCondition := resetRising AND (NOT runRequest) AND pressureValid
                  AND (pressure <= 4200.0);

// 跳闸条件
tripCondition := (runRequest AND NOT pressureValid)
                 OR (runRequest AND pressureValid AND pressure >= 4500.0);

// 更新跳闸自保持与线索足迹累积
IF resetCondition THEN
    tripLatched := FALSE;
    latchedCauseMask := 0;
ELSE
    IF tripCondition THEN
        tripLatched := TRUE;
    END_IF;
    IF tripLatched THEN
        latchedCauseMask := latchedCauseMask OR currentCauseMask;
    END_IF;
END_IF;

// 输出计算
fuelPermit := runRequest AND (NOT tripLatched);
diagnosticActive := (currentCauseMask <> 0);

// 更新历史状态
resetBtnPrev := resetBtn;

END_FUNCTION_BLOCK

(* ---- self-hard-07.st ---- *)
FUNCTION_BLOCK FB
VAR_INPUT
    mode : INT;
    resetBtn : BOOL;
    scanSeconds : REAL;
    tempSP : REAL;
    tempPV : REAL;
    flowPV : REAL;
    manualFlowSP : REAL;
    manualValve : REAL;
END_VAR
VAR_OUTPUT
    flowSP : REAL;
    valveCommand : REAL;
    fault : BOOL;
    normalMode : BOOL;
END_VAR
VAR
    firstScan : BOOL := TRUE;
    prevResetBtn : BOOL := FALSE;
    lastMode : INT := 0;
    lastFlowSP : REAL := 0.0;
    lastValveCommand : REAL := 0.0;
    iT : REAL := 0.0;
    iF : REAL := 0.0;
    eT : REAL := 0.0;
    eF : REAL := 0.0;
END_VAR

fault := (mode < 0) OR (mode > 2) OR (scanSeconds <= 0.0) OR (scanSeconds > 10.0);

IF firstScan THEN
    flowSP := manualFlowSP;
    valveCommand := manualValve;
    iT := flowSP - 1.0 * (tempSP - tempPV);
    iF := valveCommand - 2.0 * (flowSP - flowPV);
    lastMode := mode;
    lastFlowSP := flowSP;
    lastValveCommand := valveCommand;
    normalMode := FALSE;
    firstScan := FALSE;
ELSIF resetBtn AND NOT prevResetBtn THEN
    flowSP := manualFlowSP;
    valveCommand := manualValve;
    iT := flowSP - 1.0 * (tempSP - tempPV);
    iF := valveCommand - 2.0 * (flowSP - flowPV);
    lastMode := mode;
    lastFlowSP := flowSP;
    lastValveCommand := valveCommand;
    normalMode := FALSE;
ELSIF fault THEN
    flowSP := manualFlowSP;
    valveCommand := manualValve;
    iT := flowSP - 1.0 * (tempSP - tempPV);
    iF := valveCommand - 2.0 * (flowSP - flowPV);
    lastMode := mode;
    lastFlowSP := flowSP;
    lastValveCommand := valveCommand;
    normalMode := FALSE;
ELSE
    IF mode <> lastMode THEN
        (* 模式切换拍：阀位保持，流量设定按目标模式处理 *)
        valveCommand := lastValveCommand;
        IF mode = 2 THEN
            flowSP := lastFlowSP;
        ELSE
            flowSP := manualFlowSP;
        END_IF
        iT := flowSP - 1.0 * (tempSP - tempPV);
        iF := valveCommand - 2.0 * (flowSP - flowPV);
        normalMode := FALSE;
        lastMode := mode;
        lastFlowSP := flowSP;
        lastValveCommand := valveCommand;
    ELSE
        (* 正常运算拍 *)
        normalMode := TRUE;
        CASE mode OF
            0:
                flowSP := manualFlowSP;
                valveCommand := manualValve;
                iT := flowSP - 1.0 * (tempSP - tempPV);
                iF := valveCommand - 2.0 * (flowSP - flowPV);
            1:
                flowSP := manualFlowSP;
                iT := flowSP - 1.0 * (tempSP - tempPV);
                eF := flowSP - flowPV;
                iF := iF + 0.5 * eF * scanSeconds;
                valveCommand := LIMIT(0.0, 2.0 * eF + iF, 100.0);
                iF := valveCommand - 2.0 * eF;
            2:
                eT := tempSP - tempPV;
                iT := iT + 0.2 * eT * scanSeconds;
                flowSP := LIMIT(0.0, 1.0 * eT + iT, 50.0);
                iT := flowSP - 1.0 * eT;
                eF := flowSP - flowPV;
                iF := iF + 0.5 * eF * scanSeconds;
                valveCommand := LIMIT(0.0, 2.0 * eF + iF, 100.0);
                iF := valveCommand - 2.0 * eF;
        END_CASE
        lastMode := mode;
        lastFlowSP := flowSP;
        lastValveCommand := valveCommand;
    END_IF
END_IF

prevResetBtn := resetBtn;

END_FUNCTION_BLOCK

(* ---- self-medium-01.st ---- *)
TYPE ST_Recipe :
STRUCT
    recipeID : INT;
    totalRatio : REAL;
    temperature : REAL;
END_STRUCT
END_TYPE

FUNCTION_BLOCK FB
VAR_INPUT
    recipe : ARRAY[1..8] OF ST_Recipe;
    selSlot : INT;
    loadCmd : BOOL;
    running : BOOL;
END_VAR
VAR_OUTPUT
    valid : BOOL;
    loadedID : INT;
END_VAR
VAR
    lastLoadCmd : BOOL := FALSE;
    memValid : BOOL := FALSE;
    memLoadedID : INT := 0;
    risingEdge : BOOL;
END_VAR

risingEdge := loadCmd AND NOT lastLoadCmd;
lastLoadCmd := loadCmd;

IF risingEdge AND NOT running THEN
    IF (selSlot < 1) OR (selSlot > 8) THEN
        memValid := FALSE;
        memLoadedID := 0;
    ELSE
        IF recipe[selSlot].recipeID = 0 THEN
            memValid := FALSE;
            memLoadedID := 0;
        ELSIF (recipe[selSlot].totalRatio < 99.0) OR (recipe[selSlot].totalRatio > 101.0) THEN
            memValid := FALSE;
            memLoadedID := 0;
        ELSIF (recipe[selSlot].temperature < 30.0) OR (recipe[selSlot].temperature > 180.0) THEN
            memValid := FALSE;
            memLoadedID := 0;
        ELSE
            memValid := TRUE;
            memLoadedID := recipe[selSlot].recipeID;
        END_IF
    END_IF
END_IF

valid := memValid;
loadedID := memLoadedID;

END_FUNCTION_BLOCK

(* ---- self-medium-02.st ---- *)
FUNCTION_BLOCK FB
VAR_INPUT
    enable : BOOL;
    rawValue : REAL;
END_VAR
VAR_OUTPUT
    filteredValue : REAL;
    windowFull : BOOL;
    sampleCount : INT;
END_VAR
VAR
    buf : ARRAY[0..7] OF REAL;
    writeIndex : INT := 0;
    count : INT := 0;
    sum : REAL;
    i : INT;
END_VAR

IF NOT enable THEN
    count := 0;
    writeIndex := 0;
    windowFull := FALSE;
    sampleCount := 0;
ELSE
    buf[writeIndex] := rawValue;
    writeIndex := (writeIndex + 1) MOD 8;

    IF count < 8 THEN
        count := count + 1;
    END_IF;

    sum := 0.0;
    IF count > 0 THEN
        FOR i := 0 TO count - 1 DO
            sum := sum + buf[i];
        END_FOR;
        filteredValue := sum / INT_TO_REAL(count);
    END_IF;

    sampleCount := count;

    IF count >= 8 THEN
        windowFull := TRUE;
    ELSE
        windowFull := FALSE;
    END_IF;
END_IF;

END_FUNCTION_BLOCK

(* ---- self-medium-03.st ---- *)
FUNCTION_BLOCK FB
VAR_INPUT
    openBtn : BOOL;
    closeBtn : BOOL;
    openLimit : BOOL;
    closeLimit : BOOL;
    obstacle : BOOL;
END_VAR
VAR_OUTPUT
    motorUp : BOOL;
    motorDown : BOOL;
    errorFlag : BOOL;
END_VAR
VAR
    state : INT := 0; (* 0=IDLE, 1=OPENING, 2=CLOSING, 3=FAULT *)
    openBtn_prev : BOOL := FALSE;
    closeBtn_prev : BOOL := FALSE;
    openBtn_rise : BOOL;
    closeBtn_rise : BOOL;
    bothPressed : BOOL;
    bothPressed_prev : BOOL := FALSE;
    reset_rise : BOOL;
END_VAR

(* 边沿检测 *)
openBtn_rise := openBtn AND NOT openBtn_prev;
closeBtn_rise := closeBtn AND NOT closeBtn_prev;
bothPressed := openBtn AND closeBtn;
reset_rise := bothPressed AND NOT bothPressed_prev;

(* 状态机 *)
CASE state OF
    0: (* IDLE *)
        motorUp := FALSE;
        motorDown := FALSE;
        errorFlag := FALSE;
        IF openBtn_rise AND NOT openLimit THEN
            state := 1; (* OPENING *)
        ELSIF closeBtn_rise AND NOT closeLimit THEN
            state := 2; (* CLOSING *)
        END_IF;

    1: (* OPENING *)
        motorDown := FALSE;
        errorFlag := FALSE;
        IF obstacle THEN
            motorUp := FALSE;
            state := 3; (* FAULT *)
            errorFlag := TRUE;
        ELSIF openLimit THEN
            motorUp := FALSE;
            state := 0; (* IDLE *)
        ELSE
            motorUp := TRUE;
        END_IF;

    2: (* CLOSING *)
        motorUp := FALSE;
        errorFlag := FALSE;
        IF obstacle THEN
            motorDown := FALSE;
            IF openLimit THEN
                motorUp := FALSE;
                state := 0; (* IDLE *)
            ELSE
                motorUp := TRUE;
                state := 1; (* OPENING *)
            END_IF;
        ELSIF closeLimit THEN
            motorDown := FALSE;
            state := 0; (* IDLE *)
        ELSE
            motorDown := TRUE;
        END_IF;

    3: (* FAULT *)
        motorUp := FALSE;
        motorDown := FALSE;
        errorFlag := TRUE;
        IF reset_rise AND NOT obstacle THEN
            errorFlag := FALSE;
            state := 0; (* 复位到IDLE *)
        END_IF;
END_CASE

(* 更新按钮历史 *)
openBtn_prev := openBtn;
closeBtn_prev := closeBtn;
bothPressed_prev := bothPressed;

END_FUNCTION_BLOCK

(* ---- self-medium-04.st ---- *)
FUNCTION_BLOCK FB
VAR_INPUT
    startBtn : BOOL;
    resetBtn : BOOL;
    doneSensor : BOOL;
    targetVol : REAL;
    flowVol : REAL;
END_VAR
VAR_OUTPUT
    valveOpen : BOOL;
    fillsToday : INT;
END_VAR
VAR
    accVol : REAL;
    fillState : INT; (* 0=IDLE, 1=FILLING, 2=WAIT_CONFIRM *)
    startR : BOOL;
    resetR : BOOL;
    prevStart : BOOL;
    prevReset : BOOL;
END_VAR

(* 边沿检测 *)
startR := startBtn AND NOT prevStart;
resetR := resetBtn AND NOT prevReset;

IF resetR THEN
    (* 复位优先 *)
    fillsToday := 0;
    valveOpen := FALSE;
    accVol := 0.0;
    fillState := 0;
ELSE
    CASE fillState OF
        0: (* IDLE *)
            valveOpen := FALSE;
            IF startR THEN
                valveOpen := TRUE;
                accVol := 0.0;
                fillState := 1;
            END_IF;

        1: (* FILLING *)
            accVol := accVol + flowVol;
            IF accVol >= targetVol THEN
                valveOpen := FALSE;
                fillState := 2;
            ELSE
                valveOpen := TRUE;
            END_IF;

        2: (* WAIT_CONFIRM *)
            valveOpen := FALSE;
            IF doneSensor THEN
                fillsToday := fillsToday + 1;
                fillState := 0;
            END_IF;
    END_CASE;
END_IF;

(* 更新历史 *)
prevStart := startBtn;
prevReset := resetBtn;

END_FUNCTION_BLOCK

(* ---- self-medium-05.st ---- *)
FUNCTION_BLOCK FB
VAR_INPUT
    enable : BOOL;
    resetBtn : BOOL;
    scanSeconds : LREAL;
    steamFlow : LREAL;
    fuelFlow : LREAL;
    steamTemp : LREAL;
    steamPressure : LREAL;
END_VAR
VAR_OUTPUT
    qualified : BOOL;
    dataFault : BOOL;
    qualifiedTon : LREAL;
    fuelTon : LREAL;
    revenue : LREAL;
    cost : LREAL;
    netProfit : LREAL;
END_VAR
VAR
    prevReset : BOOL := FALSE;
    accQualifiedTon : LREAL := 0.0;
    accFuelTon : LREAL := 0.0;
    resetEdge : BOOL;
    canAccumulate : BOOL;
END_VAR

qualified := (steamTemp >= 447.0) AND (steamTemp <= 453.0) AND (steamPressure >= 3750.0) AND (steamPressure <= 3850.0);

dataFault := (scanSeconds <= 0.0) OR (scanSeconds > 10.0) OR (steamFlow < 0.0) OR (steamFlow > 90.0) OR (fuelFlow < 0.0) OR (fuelFlow > 6.0);

resetEdge := resetBtn AND (NOT prevReset);
prevReset := resetBtn;

IF resetEdge THEN
    accQualifiedTon := 0.0;
    accFuelTon := 0.0;
ELSE
    canAccumulate := enable AND (NOT dataFault);
    IF canAccumulate THEN
        accFuelTon := accFuelTon + (fuelFlow * scanSeconds / 1000.0);
        IF qualified THEN
            accQualifiedTon := accQualifiedTon + (steamFlow * scanSeconds / 1000.0);
        END_IF
    END_IF
END_IF

qualifiedTon := accQualifiedTon;
fuelTon := accFuelTon;
revenue := accQualifiedTon * 280.0;
cost := accFuelTon * 1500.0;
netProfit := revenue - cost;
END_FUNCTION_BLOCK

(* ---- self-medium-06.st ---- *)
FUNCTION_BLOCK FB
VAR_INPUT
    enable : BOOL;
    resetBtn : BOOL;
    sensorValid : BOOL;
    setpoint : REAL;
    temperature : REAL;
    scanSeconds : REAL;
    bias : REAL;
END_VAR
VAR_OUTPUT
    power : REAL;
    correction : REAL;
    fault : BOOL;
END_VAR
VAR
    resetPrev : BOOL;
    ePrev : REAL;
    hasHistory : BOOL;
    e : REAL;
    de : REAL;
    x : REAL;
    y : REAL;
    muNX : REAL;
    muZX : REAL;
    muPX : REAL;
    muNY : REAL;
    muZY : REAL;
    muPY : REAL;
    wNN : REAL;
    wNZ : REAL;
    wNP : REAL;
    wZN : REAL;
    wZZ : REAL;
    wZP : REAL;
    wPN : REAL;
    wPZ : REAL;
    wPP : REAL;
    sumW : REAL;
    sumWC : REAL;
    resetRising : BOOL;
    clearHistory : BOOL;
END_VAR

fault := NOT sensorValid OR scanSeconds <= 0.0 OR scanSeconds > 10.0;
resetRising := resetBtn AND NOT resetPrev;
clearHistory := NOT enable OR fault OR resetRising;

IF clearHistory THEN
    power := 0.0;
    correction := 0.0;
    ePrev := 0.0;
    hasHistory := FALSE;
ELSE
    e := setpoint - temperature;
    IF hasHistory THEN
        de := (e - ePrev) / scanSeconds;
    ELSE
        de := 0.0;
    END_IF

    x := e / 10.0;
    IF x < -1.0 THEN
        x := -1.0;
    ELSIF x > 1.0 THEN
        x := 1.0;
    END_IF

    y := de / 2.0;
    IF y < -1.0 THEN
        y := -1.0;
    ELSIF y > 1.0 THEN
        y := 1.0;
    END_IF

    IF x < 0.0 THEN
        muNX := -x;
    ELSE
        muNX := 0.0;
    END_IF
    muZX := 1.0 - ABS(x);
    IF x > 0.0 THEN
        muPX := x;
    ELSE
        muPX := 0.0;
    END_IF

    IF y < 0.0 THEN
        muNY := -y;
    ELSE
        muNY := 0.0;
    END_IF
    muZY := 1.0 - ABS(y);
    IF y > 0.0 THEN
        muPY := y;
    ELSE
        muPY := 0.0;
    END_IF

    wNN := muNX * muNY;
    wNZ := muNX * muZY;
    wNP := muNX * muPY;
    wZN := muZX * muNY;
    wZZ := muZX * muZY;
    wZP := muZX * muPY;
    wPN := muPX * muNY;
    wPZ := muPX * muZY;
    wPP := muPX * muPY;

    sumW := wNN + wNZ + wNP + wZN + wZZ + wZP + wPN + wPZ + wPP;
    IF sumW > 0.0 THEN
        sumWC := wNN * (-30.0) + wNZ * (-20.0) + wNP * (-10.0)
               + wZN * (-10.0) + wZZ * 0.0 + wZP * 10.0
               + wPN * 10.0 + wPZ * 20.0 + wPP * 30.0;
        correction := sumWC / sumW;
    ELSE
        correction := 0.0;
    END_IF

    IF correction < -30.0 THEN
        correction := -30.0;
    ELSIF correction > 30.0 THEN
        correction := 30.0;
    END_IF

    power := bias + correction;
    IF power < 0.0 THEN
        power := 0.0;
    ELSIF power > 100.0 THEN
        power := 100.0;
    END_IF

    ePrev := e;
    hasHistory := TRUE;
END_IF

resetPrev := resetBtn;
END_FUNCTION_BLOCK
